// TIA Portal V18 export
FUNCTION_BLOCK "FB_Filler"   // FB3, LAD
   VAR
      Running : Bool;   // Filler running
      Fill_Tmr : TON_TIME;
      Fill_Count : Int;   // Bottles filled
   END_VAR
BEGIN

REGION Network 1: Run latch
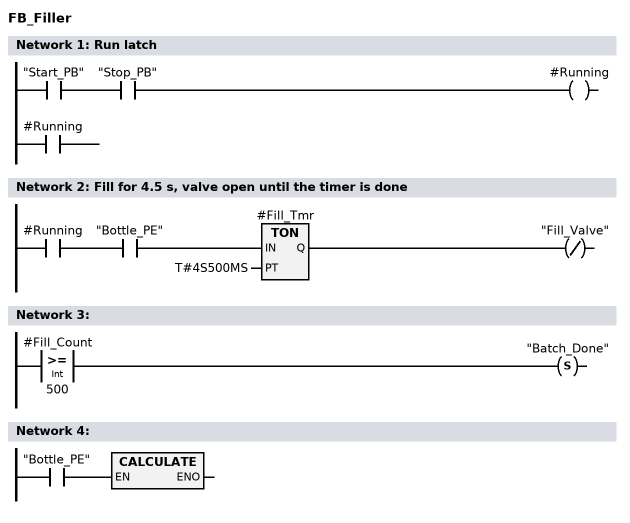
   #Running := "Start_PB" AND "Stop_PB";
END_REGION

REGION Network 2: Fill for 4.5 s, valve open until the timer is done
   RUNG wire#powerrail
      Contact( #Running )
      Contact( "Bottle_PE" )
      #Fill_Tmr.TON(pt := T#4S500MS)
      I_Coil( "Fill_Valve" )
   END_RUNG
   // the same network as SCL:
   #Fill_Tmr(IN := #Running AND "Bottle_PE", PT := T#4S500MS);   // TON
   "Fill_Valve" := NOT #Fill_Tmr.Q;
END_REGION

REGION Network 3
   RUNG wire#powerrail
      { S7_Templates := "SrcType := Int" } GE_Contact(in1 := #Fill_Count, in2 := 500)
      S_Coil( "Batch_Done" )
   END_RUNG
   // the same network as SCL:
   IF #Fill_Count >= 500 THEN "Batch_Done" := TRUE; END_IF;
END_REGION

REGION Network 4
   IF "Bottle_PE" THEN Calculate(); END_IF;
END_REGION

REGION Network 5 (SCL)
   #Fill_Count
END_REGION
END_FUNCTION_BLOCK
